Fanuc KAREL source: KO00003.KL

PROGRAM KO00003
%NOLOCKGROUP
VAR
  P1: POSITION
  P2: POSITION
  P3: POSITION
  OUT: XYZWPREXT
BEGIN
  OUT = FRAME(P1, P2, P3)
END KO00003
